// TIA Portal V21 export
// export: Created 2026-11-10T19:21:32.1837462Z, ExportSetting WithDefaults, DisplayName Totally Integrated Automation Portal, DisplayVersion V21 Update 3, DisplayName STEP 7 Professional, DisplayVersion V21 Update 3, DisplayName STEP 7 Safety, DisplayVersion V21, DisplayName Tech WebApplication, DisplayVersion V21, DisplayName WinCC Basic/Comfort/Advanced, DisplayVersion V21 Update 3, DisplayName WinCC Unified, DisplayVersion V21 Update 3
FUNCTION_BLOCK "FB_Lad_mb008"   // FB8, LAD
{ S7_Optimized_Access := 'TRUE' }
VERSION : 0.1
// stored: AutoNumber true, IsIECCheckEnabled false, IsRetainMemResEnabled false, MemoryReserve 100, SetENOAutomatically false, UDAEnableTagReadback false
   VAR_INPUT
      v_mb_addr : USInt;
   END_VAR
   VAR_OUTPUT
      v_ndr : Bool;
      v_dr : Bool;
      v_error : Bool;
      v_status : Word;
   END_VAR
   VAR_IN_OUT
      v_mb_hold_reg : Variant;
   END_VAR
   VAR
      inst { S7_SetPoint := 'True'} : Modbus_Slave;
   END_VAR
BEGIN

REGION Network 1: Description of MB_SLAVE
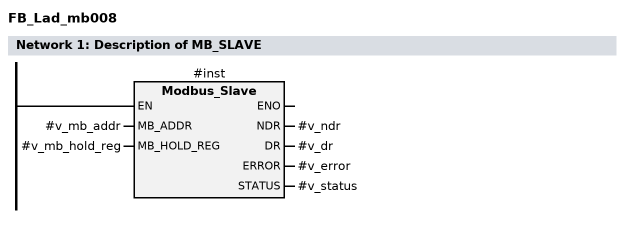
   RUNG wire#powerrail
      #inst.Modbus_Slave(MB_ADDR := #v_mb_addr, NDR => #v_ndr, DR => #v_dr, ERROR => #v_error, STATUS => #v_status, MB_HOLD_REG := #v_mb_hold_reg)
   END_RUNG
   // the same network as SCL:
   #inst(MB_ADDR := #v_mb_addr,   // Modbus_Slave
         MB_HOLD_REG := #v_mb_hold_reg,
         NDR => #v_ndr,
         DR => #v_dr,
         ERROR => #v_error,
         STATUS => #v_status);
END_REGION
END_FUNCTION_BLOCK
